(* IEC 61131-3 sources: volt/packages/volt-lsp-iec/test-corpus/bakon-nano/Device/Plc Logic/Application/Library Manager/VisuShared, 19 files *)

(* ---- EVENTPARAMSYNCFILETRANSFER.dut ---- *)
TYPE EVENTPARAMSYNCFILETRANSFER :
STRUCT
	PSAPPLICATIONNAME : POINTER TO STRING;
	UITYPE : UINT;
END_STRUCT
END_TYPE

(* ---- VISUENUMDATETIMELIBRARY.dut ---- *)
TYPE VISUENUMDATETIMELIBRARY :
(
	USESYSTIMERTC := 0,
	USEUTILSTIME := 1
);
END_TYPE

(* ---- EVENT_SYNC_FILE.gvl ---- *)
VAR_GLOBAL
	EVT_SYNCFILETRANSFER : UDINT := 16#10002;
	CMPID_CMPFILETRANSFER : UDINT := 16#5E;
	SYNCFILE_TYPE_START : UINT := 1;
	SYNCFILE_TYPE_END : UINT := 2;
END_VAR

(* ---- VISUSHARED_GLOBALS.gvl ---- *)
VAR_GLOBAL
	G_SYNCFILETRANSFEREVENT : Visu_FbSyncFileTransferEvent;
	G_UILOADTEXTLIST : UDINT;
	G_UILOADTEXTLISTOCBIT : UDINT := 0;
	G_UILOADTEXTLISTBEFOREOCBIT : UDINT := 1;
	G_UILOADTEXTLISTDLBIT : UDINT := 2;
	G_DATETIMEPROVIDER : Visu_FbDateTimeProvider;
END_VAR

(* ---- ICALLONINITIALIZEBASE.itf ---- *)
INTERFACE ICALLONINITIALIZEBASE
END_INTERFACE

METHOD INIT : BOOL
END_METHOD

(* ---- CONVERTDATETIME.pou ---- *)
FUNCTION CONVERTDATETIME : ULINT
VAR_INPUT
	UIYEAR : YEAR;
END_VAR
VAR_OUTPUT
	EERRORID : ERROR;
END_VAR
VAR_IN_OUT
	DTDATETIME : DateTime;
END_VAR
END_FUNCTION

(* ---- EXTRACTYEARMONTHDAY.pou ---- *)
FUNCTION EXTRACTYEARMONTHDAY : ERROR
VAR_INPUT
	ULIDATETIME : ULINT;
END_VAR
VAR_OUTPUT
	UIYEAR : YEAR;
	UIMONTH : MONTH;
	UIDAY : DAY;
END_VAR
END_FUNCTION

(* ---- GETLIBVERSION.pou ---- *)
FUNCTION GETLIBVERSION : VERSION
END_FUNCTION

(* ---- GETLIBVERSIONNUMBER.pou ---- *)
FUNCTION GETLIBVERSIONNUMBER : DWORD
END_FUNCTION

(* ---- GETTASKBYNAME.pou ---- *)
FUNCTION GETTASKBYNAME : BOOL
VAR_INPUT
	SZAPPNAME : STRING(CmpApp.GlobalConstants.MAX_LEN_APPLNAME);
	SZTASK : POINTER TO STRING;
END_VAR
VAR_OUTPUT
	HTASK : RTS_IEC_HANDLE;
END_VAR
END_FUNCTION

(* ---- ISLIBRELEASED.pou ---- *)
FUNCTION ISLIBRELEASED : BOOL
END_FUNCTION

(* ---- ISTASKRUNNING.pou ---- *)
FUNCTION ISTASKRUNNING : BOOL
VAR_INPUT
	HTASK : RTS_IEC_HANDLE;
	SZAPPNAME : STRING(CmpApp.GlobalConstants.MAX_LEN_APPLNAME);
END_VAR
END_FUNCTION

(* ---- LEAPYEARS.pou ---- *)
FUNCTION LEAPYEARS : UINT
VAR_INPUT
	UISTARTYEAR : YEAR;
	UIENDYEAR : YEAR;
END_VAR
VAR_OUTPUT
	EERRORID : ERROR;
END_VAR
END_FUNCTION

(* ---- LOADTEXTLISTBEFOREONLINECHANGE.pou ---- *)
FUNCTION LOADTEXTLISTBEFOREONLINECHANGE : BOOL
END_FUNCTION

(* ---- RELOADTEXTLISTSIFNECESSARY.pou ---- *)
FUNCTION RELOADTEXTLISTSIFNECESSARY : BOOL
VAR_INPUT
	BDOWNLOAD : BOOL;
	BFORCE : BOOL;
END_VAR
END_FUNCTION

(* ---- UTILTIMEZONELOCALTOUTC.pou ---- *)
FUNCTION UTILTIMEZONELOCALTOUTC : SYSTIME
VAR_INPUT
	ULILOCALTIME : SYSTIME;
END_VAR
VAR_OUTPUT
	EERRORID : ERROR;
	EPERIOD : PERIOD;
END_VAR
VAR_IN_OUT
	TZTIMEZONE : TimeZone;
END_VAR
END_FUNCTION

(* ---- VISU_FBDATETIMEPROVIDER.pou ---- *)
FUNCTION_BLOCK VISU_FBDATETIMEPROVIDER
VAR_INPUT
	ENDATETIMELIBRARY : VisuEnumDateTimeLibrary := VisuEnumDateTimeLibrary.UseSysTimeRTC;
	TZTIMEZONE : Util.TimeZone;
END_VAR
END_FUNCTION_BLOCK

METHOD CONVERTLOCALTOUTCTIME : SYSTIME
VAR_INPUT
	LOCALTIME : SYSTIME;
END_VAR
VAR_OUTPUT
	EERRORID : ERROR;
	IUTCOFFSET : INT;
END_VAR
END_METHOD

METHOD CONVERTUTCTOLOCALTIME : SYSTIME
VAR_INPUT
	UTCTIME : SYSTIME;
END_VAR
VAR_OUTPUT
	EERRORID : ERROR;
	IUTCOFFSET : INT;
END_VAR
END_METHOD

METHOD GETCURRENTLOCALTIME : SYSTIME
VAR_OUTPUT
	EERRORID : ERROR;
	IUTCOFFSET : INT;
END_VAR
END_METHOD

METHOD GETCURRENTUTCTIME : SYSTIME
VAR_OUTPUT
	EERRORID : ERROR;
END_VAR
END_METHOD

(* ---- VISU_FBINITONSTARTUP.pou ---- *)
FUNCTION_BLOCK VISU_FBINITONSTARTUP
VAR
	_ARR : ARRAY [0..(MAX_STARTUPINITIALZATIONS - 1)] OF ICallOnInitializeBase;
	_ICOUNT : INT;
	MAX_STARTUPINITIALZATIONS : INT := 5;
END_VAR
END_FUNCTION_BLOCK

METHOD CALLINITIALIZE
END_METHOD

METHOD REGISTER : BOOL
VAR_INPUT
	INSTANCE : ICallOnInitializeBase;
END_VAR
END_METHOD

(* ---- VISU_FBSYNCFILETRANSFEREVENT.pou ---- *)
FUNCTION_BLOCK VISU_FBSYNCFILETRANSFEREVENT
VAR
	_HEVENTSTART : SysTypes.RTS_IEC_HANDLE := SysTypes.RTS_INVALID_HANDLE;
	_HINTERFACESTART : SysTypes.RTS_IEC_HANDLE := SysTypes.RTS_INVALID_HANDLE;
	_ITFEVENTCALLBACK : CmpEventMgr_Interfaces.ICmpEventCallback;
END_VAR
END_FUNCTION_BLOCK

METHOD EVENTCALLBACK : SysTypes.RTS_IEC_RESULT
VAR_INPUT
	PEVENTPARAM : POINTER TO EventParam;
END_VAR
END_METHOD

METHOD FB_EXIT : BOOL
VAR_INPUT
	BINCOPYCODE : BOOL;
END_VAR
END_METHOD

METHOD FB_INIT : BOOL
VAR_INPUT
	BINITRETAINS : BOOL;
	BINCOPYCODE : BOOL;
END_VAR
END_METHOD
